Fanuc KAREL source: KA00045.KL

PROGRAM KA00045
%NOLOCKGROUP
VAR
  SRC: STRING[80]
  DST: VECTOR
BEGIN
  SRC = 'A'
  DST = SRC
END KA00045
